(* IEC 61131-3 sources: plc-ci-toolkit/src/POUs/F_Clamp, 2 files *)

(* ---- F_Clamp.decl.st ---- *)
// Назначение: ограничение значения отрезком между двумя границами.
//             Если rLow > rHigh, границы меняются местами: результат всегда лежит
//             между двумя заданными границами и не зависит от порядка аргументов.
//             NaN на входе не обрабатывается — достоверность проверяется до вызова.
// Автор:      kr0nsch
// Версия:     0.1.0
// Документ:   docs/ASSUMPTIONS.md, раздел «Семантика F_Clamp»
FUNCTION F_Clamp : REAL
VAR_INPUT
    rValue : REAL;      // ограничиваемое значение
    rLow : REAL;        // нижняя граница
    rHigh : REAL;       // верхняя граница
END_VAR
VAR
    rMin : REAL;        // нижняя граница после упорядочивания
    rMax : REAL;        // верхняя граница после упорядочивания
END_VAR

(* ---- F_Clamp.impl.st ---- *)
// Упорядочиваем границы: при rLow > rHigh меняем их местами
IF rLow <= rHigh THEN
    rMin := rLow;
    rMax := rHigh;
ELSE
    rMin := rHigh;
    rMax := rLow;
END_IF

// Ограничиваем значение; на границе возвращается сама граница
IF rValue < rMin THEN
    F_Clamp := rMin;
ELSIF rValue > rMax THEN
    F_Clamp := rMax;
ELSE
    F_Clamp := rValue;
END_IF
